(* IEC 61131-3 sources: krc-sample-programs/clamp-station-codesys/source/03_States, 2 files *)

(* ---- E_Step.st ---- *)
// The steps, a thousand apart, so steps inside a state can be added later without renumbering.
TYPE E_Step :
(
	S0_IDLE      :=    0,	// Idle: powered up and at rest. Goes straight to Not Ready
	S1_NOT_READY := 1000,	// Not Ready: waiting for the clamp to read open, both hands off, Stop not pressed
	S2_RESET     := 2000,	// Reset: clears a fault, waits for Reset to be released
	S3_READY     := 3000,	// Ready: waiting for both hand buttons
	S4_CLAMPING  := 4000,	// Clamping: valve on, setpoint out, waiting for pressure
	S5_OPENING   := 5000,	// Opening: valve off, waiting for the clamp to read open
	S6_FAULT     := 6000 	// Fault: waiting for Reset
) INT;
END_TYPE

(* ---- CONSTANTS.st ---- *)
// Named numbers the program uses, so no bare number appears in the logic.
VAR_GLOBAL CONSTANT
	AI_FULL_SCALE    : REAL := 32760.0;	// CC100 analog input raw count at 10 V (WAGO manual, section 9.4)
	AO_FULL_SCALE    : REAL := 32767.0;	// CC100 analog output raw count for 10 V (WAGO manual, section 9.4)
	PRESSURE_RANGE   : REAL := 100.0;	// psi at 10 V, for the sensor and the regulator
	PRESSURE_BAND    : REAL := 2.0;	// psi: within this much of the setpoint counts as at pressure
END_VAR
